Staubli VAL3: insertAction.pgx

public program insertAction(string x_sKey, num x_nIndex, num x_nValue, bool& x_bToSave)
  local num l_i
begin
  // insert(trajTemp:tTrajItem[x_sKey].pPointItem[x_nIndex+1])
  append(trajTemp:tTrajItem[x_sKey].pPointItem)

  for l_i = (size(trajTemp:tTrajItem[x_sKey].pPointItem)-1) to(x_nIndex+1) step -1
    //logMsg(toString("",l_i))
    call copyPoint3(x_sKey,l_i,l_i-1)
  endFor
  trajTemp:tTrajItem[x_sKey].pPointItem[x_nIndex+1].pParaItem.nMoveType=10
  trajTemp:tTrajItem[x_sKey].pPointItem[x_nIndex+1].pParaItem.nSigValue=x_nValue
  //trajTemp:libSave()
  x_bToSave=true
end
